FUNCTION_BLOCK Eject (* Composite Function Block Type *)
  (* Standard: 61499-2 *)
  (* Version 0.0, 7/2/2026, template *)
  PACKAGE Main;
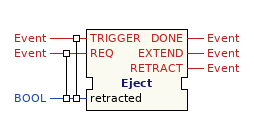
  EVENT_INPUT
    TRIGGER WITH retracted; (* Initialization Request *)
    REQ WITH retracted; (* Normal Execution Request *)
  END_EVENT
  EVENT_OUTPUT
    DONE; (* Initialization Confirm *)
    EXTEND; (* Execution Confirmation *)
    RETRACT;
  END_EVENT
  VAR_INPUT
    retracted : BOOL; (* Input event qualifier *)
  END_VAR
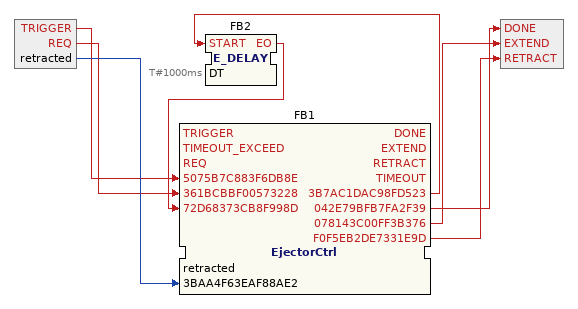
  FBS
    FB1 : EjectorCtrl;
    FB2 : E_DELAY(DT := T#1000ms);
  END_FBS
  EVENT_CONNECTIONS
    TRIGGER TO FB1.5075B7C883F6DB8E;
    REQ TO FB1.361BCBBF00573228;
    FB2.EO TO FB1.72D68373CB8F998D;
    FB1.3B7AC1DAC98FD523 TO FB2.START;
    FB1.042E79BFB7FA2F39 TO DONE;
    FB1.078143C00FF3B376 TO EXTEND;
    FB1.F0F5EB2DE7331E9D TO RETRACT;
  END_CONNECTIONS
  DATA_CONNECTIONS
    retracted TO FB1.3BAA4F63EAF88AE2;
  END_CONNECTIONS
END_FUNCTION_BLOCK
